(* IEC 61131-3 sources: plcassist-cli/packages/volt-lsp-iec/test-corpus/lenze-mid/Device/Plc Logic/Application/Library Manager/SysTimeRtc, 19 files *)

(* ---- GVL.gvl ---- *)
VAR_GLOBAL
	RTC_12HOURS : DINT := 0;
	RTC_24HOURS : DINT := 1;
	RTC_BATTERY_FAILED : DINT := 0;
	RTC_BATTERY_OK : DINT := 1;
	RTC_CTRL_CHECKBATTERY : DWORD := 0;
	RTC_CTRL_HOURMODE : DWORD := 1;
END_VAR

(* ---- SYSTIMEGETDATE.fun ---- *)
FUNCTION SYSTIMEGETDATE : UDINT
VAR_IN_OUT
	TIMEDATE : SYSTIMEDATE;
END_VAR
END_FUNCTION

(* ---- SYSTIMEGETTIMESTAMP.fun ---- *)
FUNCTION SYSTIMEGETTIMESTAMP : UDINT
END_FUNCTION

(* ---- SYSTIMERTCCONTROL.fun ---- *)
FUNCTION SYSTIMERTCCONTROL : RTS_IEC_RESULT
VAR_INPUT
	ICONTROLTAG : DINT;
END_VAR
VAR_IN_OUT
	PDICONTROLRESULT : DINT;
END_VAR
END_FUNCTION

(* ---- SYSTIMERTCCONVERTDATETOHIGHRES.fun ---- *)
FUNCTION SYSTIMERTCCONVERTDATETOHIGHRES : RTS_IEC_RESULT
VAR_IN_OUT
	PDATE : SYSTIMEDATE;
	PTIMESTAMP : SYSTIME;
END_VAR
END_FUNCTION

(* ---- SYSTIMERTCCONVERTDATETOUTC.fun ---- *)
FUNCTION SYSTIMERTCCONVERTDATETOUTC : RTS_IEC_RESULT
VAR_IN_OUT
	PDATE : SYSTIMEDATE;
	PDWTIMESTAMPUTC : DWORD;
END_VAR
END_FUNCTION

(* ---- SYSTIMERTCCONVERTHIGHRESTODATE.fun ---- *)
FUNCTION SYSTIMERTCCONVERTHIGHRESTODATE : RTS_IEC_RESULT
VAR_IN_OUT
	PTIMESTAMP : SYSTIME;
	PDATE : SYSTIMEDATE;
END_VAR
END_FUNCTION

(* ---- SYSTIMERTCCONVERTHIGHRESTOLOCAL.fun ---- *)
FUNCTION SYSTIMERTCCONVERTHIGHRESTOLOCAL : RTS_IEC_RESULT
VAR_IN_OUT
	PTIMESTAMP : SYSTIME;
	PDATE : SYSTIMEDATE;
END_VAR
END_FUNCTION

(* ---- SYSTIMERTCCONVERTLOCALTOHIGHRES.fun ---- *)
FUNCTION SYSTIMERTCCONVERTLOCALTOHIGHRES : RTS_IEC_RESULT
VAR_IN_OUT
	PDATE : SYSTIMEDATE;
	PTIMESTAMP : SYSTIME;
END_VAR
END_FUNCTION

(* ---- SYSTIMERTCCONVERTLOCALTOUTC.fun ---- *)
FUNCTION SYSTIMERTCCONVERTLOCALTOUTC : RTS_IEC_RESULT
VAR_INPUT
	DWTIMESTAMPLOCAL : DWORD;
END_VAR
VAR_IN_OUT
	PDWTIMESTAMPUTC : DWORD;
END_VAR
END_FUNCTION

(* ---- SYSTIMERTCCONVERTUTCTODATE.fun ---- *)
FUNCTION SYSTIMERTCCONVERTUTCTODATE : RTS_IEC_RESULT
VAR_INPUT
	DWTIMESTAMPUTC : DWORD;
END_VAR
VAR_IN_OUT
	PDATE : SYSTIMEDATE;
END_VAR
END_FUNCTION

(* ---- SYSTIMERTCCONVERTUTCTOLOCAL.fun ---- *)
FUNCTION SYSTIMERTCCONVERTUTCTOLOCAL : RTS_IEC_RESULT
VAR_INPUT
	DWTIMESTAMPUTC : DWORD;
END_VAR
VAR_IN_OUT
	PDWTIMESTAMPLOCAL : DWORD;
END_VAR
END_FUNCTION

(* ---- SYSTIMERTCGET.fun ---- *)
FUNCTION SYSTIMERTCGET : DWORD
VAR_IN_OUT
	PRESULT : RTS_IEC_RESULT;
END_VAR
END_FUNCTION

(* ---- SYSTIMERTCGETTIMEZONE.fun ---- *)
FUNCTION SYSTIMERTCGETTIMEZONE : RTS_IEC_RESULT
VAR_IN_OUT
	PTIMEZONE : TimezoneInformation;
END_VAR
END_FUNCTION

(* ---- SYSTIMERTCGETTIMEZONE2.fun ---- *)
FUNCTION SYSTIMERTCGETTIMEZONE2 : RTS_IEC_RESULT
VAR_IN_OUT
	PTZI : TimezoneInformation2;
END_VAR
END_FUNCTION

(* ---- SYSTIMERTCHIGHRESGET.fun ---- *)
FUNCTION SYSTIMERTCHIGHRESGET : RTS_IEC_RESULT
VAR_IN_OUT
	PTIMESTAMP : SYSTIME;
END_VAR
END_FUNCTION

(* ---- SYSTIMERTCHIGHRESSET.fun ---- *)
FUNCTION SYSTIMERTCHIGHRESSET : RTS_IEC_RESULT
VAR_IN_OUT
	PTIMESTAMP : SYSTIME;
END_VAR
END_FUNCTION

(* ---- SYSTIMERTCSET.fun ---- *)
FUNCTION SYSTIMERTCSET : RTS_IEC_RESULT
VAR_INPUT
	ULTIMESTAMP : DWORD;
END_VAR
END_FUNCTION

(* ---- SYSTIMERTCSETTIMEZONE.fun ---- *)
FUNCTION SYSTIMERTCSETTIMEZONE : RTS_IEC_RESULT
VAR_IN_OUT
	PTIMEZONE : TimezoneInformation;
END_VAR
END_FUNCTION
